Fanuc KAREL source: KA00118.KL

PROGRAM KA00118
%NOLOCKGROUP
VAR
  SRC: CONFIG
  DST: CONFIG
BEGIN
  SRC.CFG_FLIP = TRUE
  DST = SRC
END KA00118
